(* Single Vertical Tank with Operator Control Panel *)

PROGRAM main
  VAR
    TLB1 AT %IX0.1 : BOOL; (* Upper Binary Tank Level Sensor *)
    TLB2 AT %IX0.2 : BOOL; (* Lower Binary Tank Level Sensor *)
    MV1 AT %QX0.1 : BOOL;
    MV2 AT %QX0.2 : BOOL; (* Outlet Valve *)
    Start AT %IX1.0 : BOOL;
    Stop AT %IX1.1 : BOOL;
    CycleOn AT %QX1.0 : BOOL; (* Simple Lamp Indicating Cycle *)
    Buzzer AT %QX1.1 : BOOL;
    SR0 : SR;
    SR1 : SR;
  END_VAR
  VAR  (* added by the conversion: wires and edge detectors of the diagram *)
    R_TRIG1 : R_TRIG;
    F_TRIG2 : F_TRIG;
  END_VAR

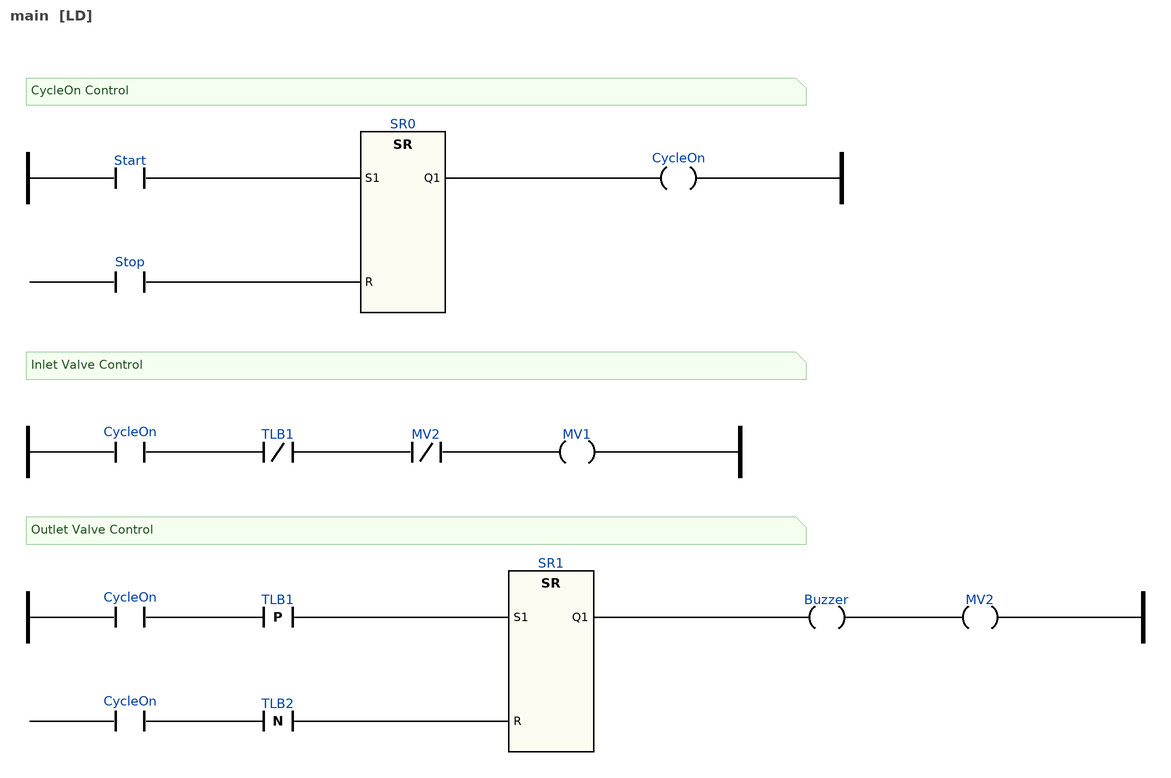
(* LD diagram, written out as Structured Text *)
(* CycleOn Control *)
SR0(S1 := Start, R := Stop);
CycleOn := SR0.Q1;
(* Inlet Valve Control *)
MV1 := CycleOn AND NOT TLB1 AND NOT MV2;
(* Outlet Valve Control *)
R_TRIG1(CLK := TLB1);
F_TRIG2(CLK := TLB2);
SR1(S1 := CycleOn AND R_TRIG1.Q, R := CycleOn AND F_TRIG2.Q);
Buzzer := SR1.Q1;
MV2 := SR1.Q1;
END_PROGRAM
